// SIMATIC S7-200 project (STEP 7-Micro/WIN), CPU 224XP CN REL 02.01

SYMBOL_TABLE USER1
PUNTERO          VD0      // PUNTERO PARA EL DATALOGGER
CONTADOR         VD4      // IGNORAR
END_SYMBOL_TABLE

SYMBOL_TABLE DATOSP1
DATO0            VD100
DATO1            VD104
DATO2            VD108
DATO3            VD112
DATO4            VD116
DATO5            VD120
DATO6            VD124
DATO7            VD128
DATO8            VD132
DATO9            VD136
DATO10           VD140
DATO11           VD144
DATO12           VD148
DATO13           VD152
DATO14           VD156
DATO15           VD160
DATO16           VD164
DATO17           VD168
DATO18           VD172
DATO19           VD176
DATO20           VD180
DATO21           VD184
DATO22           VD188
DATO23           VD192
DATO24           VD196
DATO25           VD200
DATO26           VD204
DATO27           VD208
DATO28           VD212
DATO29           VD216
DATO30           VD220
DATO31           VD224
DATO32           VD228
DATO33           VD232
DATO34           VD236
DATO35           VD240
DATO36           VD244
DATO37           VD248
DATO38           VD252
DATO39           VD256
DATO40           VD260
DATO41           VD264
DATO42           VD268
DATO43           VD272
DATO44           VD276
DATO45           VD280
DATO46           VD284
DATO47           VD288
DATO48           VD292
DATO49           VD296
DATO50           VD300
DATO51           VD304
DATO52           VD308
DATO53           VD312
DATO54           VD316
DATO55           VD320
DATO56           VD324
DATO57           VD328
DATO58           VD332
DATO59           VD336
DATO60           VD340
DATO61           VD344
DATO62           VD348
DATO63           VD352
DATO64           VD356
DATO65           VD360
DATO66           VD364
DATO67           VD368
DATO68           VD372
DATO69           VD376
DATO70           VD380
DATO71           VD384
DATO72           VD388
DATO73           VD392
DATO74           VD396
DATO75           VD400
DATO76           VD404
DATO77           VD408
DATO78           VD412
DATO79           VD416
DATO80           VD420
DATO81           VD424
DATO82           VD428
DATO83           VD432
DATO84           VD436
DATO85           VD440
DATO86           VD444
DATO87           VD448
DATO88           VD452
DATO89           VD456
DATO90           VD460
DATO91           VD464
DATO92           VD468
DATO93           VD472
DATO94           VD476
DATO95           VD480
DATO96           VD484
DATO97           VD488
DATO98           VD492
DATO99           VD496
DATO100          VD500
DATO101          VD504
DATO102          VD508
DATO103          VD512
DATO104          VD516
DATO105          VD520
DATO106          VD524
DATO107          VD528
DATO108          VD532
DATO109          VD536
DATO110          VD540
DATO111          VD544
DATO112          VD548
DATO113          VD552
DATO114          VD556
DATO115          VD560
DATO116          VD564
DATO117          VD568
DATO118          VD572
DATO119          VD576
DATO120          VD580
DATO121          VD584
DATO122          VD588
DATO123          VD592
DATO124          VD596
DATO125          VD600
DATO126          VD604
DATO127          VD608
DATO128          VD612
DATO129          VD616
DATO130          VD620
DATO131          VD624
DATO132          VD628
DATO133          VD632
DATO134          VD636
DATO135          VD640
DATO136          VD644
DATO137          VD648
DATO138          VD652
DATO139          VD656
DATO140          VD660
DATO141          VD664
DATO142          VD668
DATO143          VD672
DATO144          VD676
DATO145          VD680
DATO146          VD684
DATO147          VD688
DATO148          VD692
DATO149          VD696
END_SYMBOL_TABLE

SYMBOL_TABLE DATOSP2
DATO150          VD700
DATO151          VD704
DATO152          VD708
DATO153          VD712
DATO154          VD716
DATO155          VD720
DATO156          VD724
DATO157          VD728
DATO158          VD732
DATO159          VD736
DATO160          VD740
DATO161          VD744
DATO162          VD748
DATO163          VD752
DATO164          VD756
DATO165          VD760
DATO166          VD764
DATO167          VD768
DATO168          VD772
DATO169          VD776
DATO170          VD780
DATO171          VD784
DATO172          VD788
DATO173          VD792
DATO174          VD796
DATO175          VD800
DATO176          VD804
DATO177          VD808
DATO178          VD812
DATO179          VD816
DATO180          VD820
DATO181          VD824
DATO182          VD828
DATO183          VD832
DATO184          VD836
DATO185          VD840
DATO186          VD844
DATO187          VD848
DATO188          VD852
DATO189          VD856
DATO190          VD860
DATO191          VD864
DATO192          VD868
DATO193          VD872
DATO194          VD876
DATO195          VD880
DATO196          VD884
DATO197          VD888
DATO198          VD892
DATO199          VD896
DATO200          VD900
DATO201          VD904
DATO202          VD908
DATO203          VD912
DATO204          VD916
DATO205          VD920
DATO206          VD924
DATO207          VD928
DATO208          VD932
DATO209          VD936
DATO210          VD940
DATO211          VD944
DATO212          VD948
DATO213          VD952
DATO214          VD956
DATO215          VD960
DATO216          VD964
DATO217          VD968
DATO218          VD972
DATO219          VD976
DATO220          VD980
DATO221          VD984
DATO222          VD988
DATO223          VD992
DATO224          VD996
DATO225          VD1000
DATO226          VD1004
DATO227          VD1008
DATO228          VD1012
DATO229          VD1016
DATO230          VD1020
DATO231          VD1024
DATO232          VD1028
DATO233          VD1032
DATO234          VD1036
DATO235          VD1040
DATO236          VD1044
DATO237          VD1048
DATO238          VD1052
DATO239          VD1056
DATO240          VD1060
DATO241          VD1064
DATO242          VD1068
DATO243          VD1072
DATO244          VD1076
DATO245          VD1080
DATO246          VD1084
DATO247          VD1088
DATO248          VD1092
DATO249          VD1096
DATO250          VD1100
DATO251          VD1104
DATO252          VD1108
DATO253          VD1112
DATO254          VD1116
DATO255          VD1120
DATO256          VD1124
DATO257          VD1128
DATO258          VD1132
DATO259          VD1136
DATO260          VD1140
DATO261          VD1144
DATO262          VD1148
DATO263          VD1152
DATO264          VD1156
DATO265          VD1160
DATO266          VD1164
DATO267          VD1168
DATO268          VD1172
DATO269          VD1176
DATO270          VD1180
DATO271          VD1184
DATO272          VD1188
DATO273          VD1192
DATO274          VD1196
DATO275          VD1200
DATO276          VD1204
DATO277          VD1208
DATO278          VD1212
DATO279          VD1216
DATO280          VD1220
DATO281          VD1224
DATO282          VD1228
DATO283          VD1232
DATO284          VD1236
DATO285          VD1240
DATO286          VD1244
DATO287          VD1248
DATO288          VD1252
DATO289          VD1256
DATO290          VD1260
DATO291          VD1264
DATO292          VD1268
DATO293          VD1272
DATO294          VD1276
DATO295          VD1280
DATO296          VD1284
DATO297          VD1288
DATO298          VD1292
DATO299          VD1296
END_SYMBOL_TABLE

SYMBOL_TABLE DATOSP3
DATO300          VD1300
DATO301          VD1304
DATO302          VD1308
DATO303          VD1312
DATO304          VD1316
DATO305          VD1320
DATO306          VD1324
DATO307          VD1328
DATO308          VD1332
DATO309          VD1336
DATO310          VD1340
DATO311          VD1344
DATO312          VD1348
DATO313          VD1352
DATO314          VD1356
DATO315          VD1360
DATO316          VD1364
DATO317          VD1368
DATO318          VD1372
DATO319          VD1376
DATO320          VD1380
DATO321          VD1384
DATO322          VD1388
DATO323          VD1392
DATO324          VD1396
DATO325          VD1400
DATO326          VD1404
DATO327          VD1408
DATO328          VD1412
DATO329          VD1416
DATO330          VD1420
DATO331          VD1424
DATO332          VD1428
DATO333          VD1432
DATO334          VD1436
DATO335          VD1440
DATO336          VD1444
DATO337          VD1448
DATO338          VD1452
DATO339          VD1456
DATO340          VD1460
DATO341          VD1464
DATO342          VD1468
DATO343          VD1472
DATO344          VD1476
DATO345          VD1480
DATO346          VD1484
DATO347          VD1488
DATO348          VD1492
DATO349          VD1496
DATO350          VD1500
DATO351          VD1504
DATO352          VD1508
DATO353          VD1512
DATO354          VD1516
DATO355          VD1520
DATO356          VD1524
DATO357          VD1528
DATO358          VD1532
DATO359          VD1536
DATO360          VD1540
DATO361          VD1544
DATO362          VD1548
DATO363          VD1552
DATO364          VD1556
DATO365          VD1560
DATO366          VD1564
DATO367          VD1568
DATO368          VD1572
DATO369          VD1576
DATO370          VD1580
DATO371          VD1584
DATO372          VD1588
DATO373          VD1592
DATO374          VD1596
DATO375          VD1600
DATO376          VD1604
DATO377          VD1608
DATO378          VD1612
DATO379          VD1616
DATO380          VD1620
DATO381          VD1624
DATO382          VD1628
DATO383          VD1632
DATO384          VD1636
DATO385          VD1640
DATO386          VD1644
DATO387          VD1648
DATO388          VD1652
DATO389          VD1656
DATO390          VD1660
DATO391          VD1664
DATO392          VD1668
DATO393          VD1672
DATO394          VD1676
DATO395          VD1680
DATO396          VD1684
DATO397          VD1688
DATO398          VD1692
DATO399          VD1696
DATO400          VD1700
DATO401          VD1704
DATO402          VD1708
DATO403          VD1712
DATO404          VD1716
DATO405          VD1720
DATO406          VD1724
DATO407          VD1728
DATO408          VD1732
DATO409          VD1736
DATO410          VD1740
DATO411          VD1744
DATO412          VD1748
DATO413          VD1752
DATO414          VD1756
DATO415          VD1760
DATO416          VD1764
DATO417          VD1768
DATO418          VD1772
DATO419          VD1776
DATO420          VD1780
DATO421          VD1784
DATO422          VD1788
DATO423          VD1792
DATO424          VD1796
DATO425          VD1800
DATO426          VD1804
DATO427          VD1808
DATO428          VD1812
DATO429          VD1816
DATO430          VD1820
DATO431          VD1824
DATO432          VD1828
DATO433          VD1832
DATO434          VD1836
DATO435          VD1840
DATO436          VD1844
DATO437          VD1848
DATO438          VD1852
DATO439          VD1856
DATO440          VD1860
DATO441          VD1864
DATO442          VD1868
DATO443          VD1872
DATO444          VD1876
DATO445          VD1880
DATO446          VD1884
DATO447          VD1888
DATO448          VD1892
DATO449          VD1896
END_SYMBOL_TABLE

SYMBOL_TABLE S7-200 Symbols
Always_On        SM0.0    // Always ON
First_Scan_On    SM0.1    // ON for the first scan cycle only
Time_0_Intrvl    SMB34    // Specifies time interval (in 1-ms increments from 5 to 255) of interrupt 0.
HSC0_Ctrl        SMB37    // Configure and control HSC0
HSC0_CV          SMD38    // HSC0 new current value
HSC0_PV          SMD42    // HSC0 new preset value
END_SYMBOL_TABLE

ORGANIZATION_BLOCK MAIN:OB1
TITLE=UNIV. HERRERA TOLA GABRIEL SEBASTIAN - ETN1034 - I/2026
// DESCRIPCIÓN GENERAL:
// Este programa realiza la adquisición de datos de posición mediante un encoder incremental acoplado a un motor trifásico. Implementa una interrupción temporizada (SMB34) para el muestreo síncrono del Contador de Alta Velocidad (HSC), almacenando los registros en un buffer de memoria V mediante direccionamiento indirecto (punteros).
// 
// LÓGICA DE CONTROL:
// 
// - Entrada I1.3 (Arranque): Activa la marcha del motor a través del variador de frecuencia y habilita el proceso de captura de datos en tiempo real.
// - Intervalo de Muestreo: 10 ms.
BEGIN
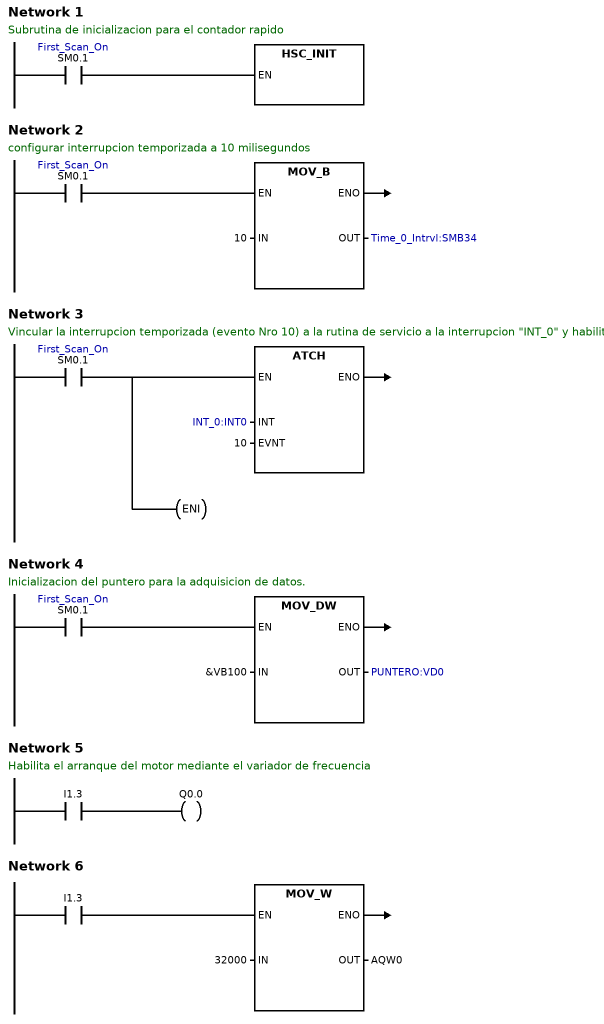
Network 1
// Subrutina de inicializacion para el contador rapido
LD     First_Scan_On:SM0.1
CALL   HSC_INIT:SBR1
Network 2
// configurar interrupcion temporizada a 10 milisegundos
LD     First_Scan_On:SM0.1
MOVB   10, Time_0_Intrvl:SMB34
Network 3
// Vincular la interrupcion temporizada (evento Nro 10) a la rutina de servicio a la interrupcion "INT_0" y habilitar las intrrupciones (ENI)
LD     First_Scan_On:SM0.1
ATCH   INT_0:INT0, 10
ENI
Network 4
// Inicializacion del puntero para la adquisicion de datos.
LD     First_Scan_On:SM0.1
MOVD   &VB100, PUNTERO:VD0
Network 5
// Habilita el arranque del motor mediante el variador de frecuencia
LD     I1.3
=      Q0.0
Network 6
LD     I1.3
MOVW   32000, AQW0
END_ORGANIZATION_BLOCK

SUBROUTINE_BLOCK HSC_INIT:SBR1
TITLE=
BEGIN
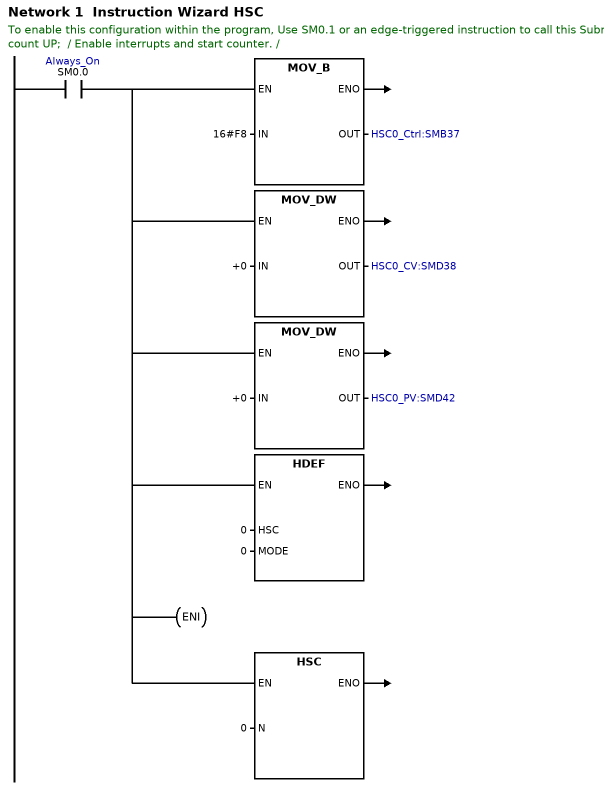
Network 1 // Instruction Wizard HSC
// To enable this configuration within the program, Use SM0.1 or an edge-triggered instruction to call this Subroutine once from the MAIN program block.  
// Configure HC0 for Mode 0; CV = 0; PV = 0; count UP; 
// Enable interrupts and start counter.
// 
//Set control bits: count UP; enabled; 
//Load CV
//Load PV
LD     Always_On:SM0.0
MOVB   16#F8, HSC0_Ctrl:SMB37
MOVD   +0, HSC0_CV:SMD38
MOVD   +0, HSC0_PV:SMD42
HDEF   0, 0
ENI
HSC    0
END_SUBROUTINE_BLOCK

INTERRUPT_BLOCK INT_0:INT0
TITLE=I1.3 ES LA ENTRADA DEL BOTON DE ARRANQUE
BEGIN
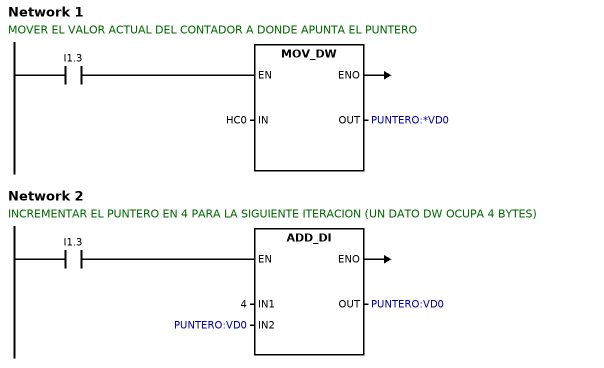
Network 1
// MOVER EL VALOR ACTUAL DEL CONTADOR A DONDE APUNTA EL PUNTERO
LD     I1.3
MOVD   HC0, *PUNTERO:VD0
Network 2
// INCREMENTAR EL PUNTERO EN 4 PARA LA SIGUIENTE ITERACION (UN DATO DW OCUPA 4 BYTES)
LD     I1.3
+D     4, PUNTERO:VD0
END_INTERRUPT_BLOCK

// (further data pages could not be read)
